(* IEC 61131-3 sources: plc-vscode/tests/st/all/trust-platform/examples/OSCAT/recipe_batch_stack/non-oop/src, 3 files *)

(* ---- Configuration.st ---- *)
CONFIGURATION RecipeBatchStackClassicConfiguration
RESOURCE Cpu0 ON PLC
    TASK MainTask (INTERVAL := T#100ms, PRIORITY := 1);
    PROGRAM Main WITH MainTask : Main;
END_RESOURCE
END_CONFIGURATION

(* ---- Main.st ---- *)
PROGRAM Main
VAR
    RecipeStack : STACK_16;
    ActiveRecipeId : DWORD;
END_VAR

RecipeStack(DIN := DWORD#16#A001, E := TRUE, RD := FALSE, WD := TRUE, RST := FALSE);
RecipeStack(DIN := DWORD#16#A002, E := TRUE, RD := FALSE, WD := TRUE, RST := FALSE);
RecipeStack(DIN := DWORD#0, E := TRUE, RD := TRUE, WD := FALSE, RST := FALSE);
ActiveRecipeId := RecipeStack.DOUT;
END_PROGRAM

(* ---- Tests.st ---- *)
TEST_PROGRAM RecipeBatchStackClassicReturnsLatestRecipe
VAR
    RecipeStack : STACK_16;
END_VAR

RecipeStack(DIN := DWORD#0, E := TRUE, RD := FALSE, WD := FALSE, RST := TRUE);
RecipeStack(DIN := DWORD#16#A001, E := TRUE, RD := FALSE, WD := TRUE, RST := FALSE);
RecipeStack(DIN := DWORD#16#A002, E := TRUE, RD := FALSE, WD := TRUE, RST := FALSE);
RecipeStack(DIN := DWORD#0, E := TRUE, RD := TRUE, WD := FALSE, RST := FALSE);

ASSERT_EQUAL(EXPECTED := DWORD#16#A002, ACTUAL := RecipeStack.DOUT);
END_TEST_PROGRAM
